(* IEC 61131-3 sources: BODAS-HelloWorld/st/bodas_rc18_12_40/plc_logic/application/02_easyconfig/easyconfig_import/bdl, 4 files *)

(* ---- bds_snsrdsa_inst_te-bds_snsrDsa_inst_te.st ---- *)
(* --- Interface --- *)
{attribute 'qualified_only' := ''}
{attribute 'strict' := ''}
TYPE bds_snsrDsa_inst_te : (
		bds_snsrDsa_numInst_E
	) USINT;
END_TYPE

(* ---- bds_snsrdst_inst_te-bds_snsrDst_inst_te.st ---- *)
(* --- Interface --- *)
{attribute 'qualified_only' := ''}
{attribute 'strict' := ''}
TYPE bds_snsrDst_inst_te : (
		SpdSnsr_E := 0,
		bds_snsrDst_numInst_E
	) USINT;
END_TYPE

(* ---- bds_snsrpal_inst_te-bds_snsrPal_inst_te.st ---- *)
(* --- Interface --- *)
{attribute 'qualified_only' := ''}
{attribute 'strict' := ''}
TYPE bds_snsrPal_inst_te : (
		bds_snsrPal_numInst_E
	) USINT;
END_TYPE

(* ---- bds_snsrpr4_inst_te-bds_snsrPr4_inst_te.st ---- *)
(* --- Interface --- *)
{attribute 'qualified_only' := ''}
{attribute 'strict' := ''}
TYPE bds_snsrPr4_inst_te : (
		pSnsr_E := 0,
		SENT_K36_E,
		SENT_K53_E,
		SENT_K57_E,
		bds_snsrPr4_numInst_E
	) USINT;
END_TYPE
